// TIA Portal V19 export
TYPE "ST_REER_INPUT"
   STRUCT
      INPUT : Array[0..32] of "ST_System_IO";
   END_STRUCT;
END_TYPE
